TYPE ST_ServiceTimeCollectionStatus :
STRUCT
	RecordCount : UINT;
	// The first records are preserved when capacity is exhausted.
	Overflow : BOOL;
	Records : ARRAY[1..Param_Config.MaxServiceTimeRecords] OF ST_ServiceStepTimeInfo;
END_STRUCT
END_TYPE

(* stored: Version 1.1.0.1, ProductVersion 3.1.4026.18
   DUT ST_ServiceTimeCollectionStatus: Id {2aeb22a5-aae2-4f9b-9e16-23f5d335838b} *)
